// TIA Portal V20 export
// export: Created 2026-10-19T18:04:33.3902132Z, ExportSetting WithDefaults, DisplayName Totally Integrated Automation Portal, DisplayVersion V20 Update 6, DisplayName TIA Portal Openness, DisplayVersion V20 Update 6, DisplayName TIA Portal Version Control Interface, DisplayVersion V20 Update 6, DisplayName SINAMICS Startdrive Advanced, DisplayVersion V20 SP1, DisplayName SINAMICS Startdrive G130, G150, S120, S150, SINAMICS MV, G220, S200, S210, DisplayVersion V20 SP1, DisplayName SINAMICS Startdrive G110M, G120, G120C, G120D, G120P, G115D, DisplayVersion V20 SP1, DisplayName STEP 7 Professional, DisplayVersion V20 Update 6, DisplayName STEP 7 Safety, DisplayVersion V20 Update 2, DisplayName WinCC Basic/Comfort/Advanced, DisplayVersion V20 Update 6, DisplayName WinCC Unified, DisplayVersion V20 Update 6
DATA_BLOCK "PopUps_DB"   // DB20
{ S7_Optimized_Access := 'TRUE' }
VERSION : 0.1
// stored: AutoNumber true, DBAccessibleFromOPCUA true, DBAccessibleFromWebserver true, IsOnlyStoredInLoadMemory false, IsRetainMemResEnabled false, IsWriteProtectedInAS false, MemoryReserve 100
   VAR
      Cnv_Select : DInt;
      Cnv_Select_Old : DInt;
      VTD_Select : DInt;
      Buffer_Cnv_Settings : "Buffer_Cnv_Settings";
      ECnv_Settings { S7_SetPoint := 'True'} : "ECnv_Settings";
      Inbound_Cnv_Settings { S7_SetPoint := 'True'} : "Inbound_Cnv_Settings";
      Outbound_Cnv_Settings { S7_SetPoint := 'True'} : "Outbound_Cnv_Settings";
      PopUp_Cnv_settings { S7_SetPoint := 'True'} : "PopUp_Cnv_Settings";
      System_Settings { S7_SetPoint := 'True'} : "System_Settings";
      VTD_Settings { S7_SetPoint := 'True'} : "VTD_Settings";
      Shuttle_MQTT_Settings { S7_SetPoint := 'True'} : "MQTT_Settings";
      LockingPins : Struct
         Faceplate : "FacePlate_LP_UDT";
         ExtendLeft { S7_SetPoint := 'True'} : Bool;
         RetractLeft { S7_SetPoint := 'True'} : Bool;
         ExtendRight { S7_SetPoint := 'True'} : Bool;
         RetractRight { S7_SetPoint := 'True'} : Bool;
         Extend_All : Bool;
         Retract_All : Bool;
      END_STRUCT;
      BSettings_Visibility : Bool;
      ESettings_Visibility : Bool;
      InSettings_Visibility : Bool;
      OutSettings_Visibility : Bool;
      PSettings_Visibility : Bool;
   END_VAR
BEGIN
   Shuttle_MQTT_Settings.MQTT_Con_Params.hwId := 64;
   Shuttle_MQTT_Settings.MQTT_Con_Params.broker := '10.0.34.2';
   Shuttle_MQTT_Settings.Client_ID := WSTRING#'PLC';
   Shuttle_MQTT_Settings.Username := WSTRING#'Devin';
   Shuttle_MQTT_Settings.Password := WSTRING#'1';
   Shuttle_MQTT_Settings.Retain := TRUE;
END_DATA_BLOCK
